(* IEC 61131-3 sources: tsplc/packages/vscode-extension/tests/fixtures/blueprint/types/ST_Reader, 3 files *)

(* ---- ST_Reader.st ---- *)
(*
Fixed-mount barcode reader EtherNet/IP signals from input assembly 11 and output assembly 21. Input is reader-to-PLC; Output is PLC-to-reader.
*)
TYPE ST_Reader :
STRUCT
	(* Reader-to-PLC signals from input assembly 11. *)
	Input : ST_ReaderInput;
	(* PLC-to-reader signals in output assembly 21. *)
	Output : ST_ReaderOutput;
END_STRUCT
END_TYPE

(* ---- ST_ReaderInput.st ---- *)
(*
Fixed-mount barcode reader EtherNet/IP signals from input assembly 11 and output assembly 21. Input is reader-to-PLC; Output is PLC-to-reader.
*)
TYPE ST_ReaderInput :
STRUCT
	(* Ready to accept an EtherNet/IP trigger; byte 0 bit 0. *)
	TriggerReady : BOOL;
	(* Acknowledges Trigger and remains set until Trigger is cleared; byte 0 bit 1. *)
	TriggerAck : BOOL;
	(* Image acquisition is in progress; byte 0 bit 2. *)
	Acquiring : BOOL;
	(* An acquisition trigger was missed; cleared by the next successful acquisition; byte 0 bit 3. *)
	MissedAcq : BOOL;
	(* Toggles for each completed decode, including no-read results; byte 1 bit 1. *)
	DecodeCompleteToggle : BOOL;
	(* A result was discarded because the results queue was full; byte 1 bit 2. *)
	ResultsBufferOverrun : BOOL;
	(* Result metadata and data are available for consumption; byte 1 bit 3. *)
	ResultsAvailable : BOOL;
	(* Reader-reported general fault indication; byte 1 bit 7. *)
	GeneralFault : BOOL;
	(* Software-event acknowledgements, bits corresponding to Output.SoftEvent; byte 2. *)
	SoftEventAck : BYTE;
	(* 16-bit identifier of the next trigger; bytes 6-7. *)
	TriggerID : UINT;
	(* Trigger identifier associated with these results; bytes 8-9. *)
	ResultID : UINT;
	(* Result flags: bit 0 read, 1 validated, 2 verified, 3 trigger overrun, 4 acquisition buffer overflow; bytes 10-11. *)
	ResultCode : WORD;
	(* Unused result extension word in the documented assembly; bytes 12-13. *)
	ResultExtended : WORD;
	(* Number of result bytes to consume from ResultData; bytes 14-15. *)
	ResultLength : UINT;
	(* Decode-result bytes, preserving the reader's configured output format; assembly bytes 16-499. *)
	ResultData : ARRAY[0..483] OF BYTE;
END_STRUCT
END_TYPE

(* ---- ST_ReaderOutput.st ---- *)
(*
Fixed-mount barcode reader EtherNet/IP signals from input assembly 11 and output assembly 21. Input is reader-to-PLC; Output is PLC-to-reader.
*)
TYPE ST_ReaderOutput :
STRUCT
	(* Enables EtherNet/IP triggering; byte 0 bit 0. *)
	TriggerEnable : BOOL;
	(* Acquisition request; hold until TriggerAck, then clear; byte 0 bit 1. *)
	Trigger : BOOL;
	(* Holds queued results until the ResultsAck handshake; byte 0 bit 2. *)
	BufferResultsEnable : BOOL;
	(* Acknowledges consumed results; clear after ResultsAvailable clears; byte 0 bit 3. *)
	ResultsAck : BOOL;
	(* Rising-edge requests: bits 0 train code, 1 train match string, 2 train focus, 3 train brightness, 4 untrain, 6 execute command, 7 set match string; bit 5 reserved. Byte 1. *)
	SoftEvent : BYTE;
	(* User-data option word from the documented assembly; bytes 4-5. *)
	UserDataOption : WORD;
	(* Number of user-data bytes supplied to the reader; bytes 6-7. *)
	UserDataLength : UINT;
	(* User-data bytes for supported operations such as reader commands and match strings; assembly bytes 8-499. *)
	UserData : ARRAY[0..491] OF BYTE;
END_STRUCT
END_TYPE
